// SIMATIC S7-200 project (STEP 7-Micro/WIN), CPU 226 CN REL 02.01

SYMBOL_TABLE USUARIO1
ANTI_HORARIO     Q0.4     // Giro del brazo en sentido antihorario
HORARIO          Q0.5     // Giro del brazo en sentido horario
CIL_DOBLE        Q0.6     // Extencion del brazo neumatico
ELEVACION        Q0.3     // Elevacion del brazo neumatico
PINZA_ABIERTA    Q1.0     // Pinza abierta del brazo neumatico
PINZA_CERRADA    Q0.7     // Pinza cerrada del brazo neumatico
DIRECCION_MOTOR  Q0.1     // Drceccion del motor (adelante o atras)
HL1              Q1.5     // Lampara de señalizacion amarilla
HL2              Q1.6     // Lampara de señaliacion verde
HL3              Q1.7     // Lampara de señalizacion roja
CIL_ABAJO        I0.3     // Sensor indicador de cilindro abajo
CIL_ARRIBA       I0.4     // Sensor indicador de cilindro arriba
CIL_EXT          I0.7     // Sensor indicador de cilindro doble extendido
CIL_RET          I1.0     // Sensor indicador de cilindro doble retraido
PINZA_CERRADO    I1.1     // Sensor indicador de Pinza cerrada
ROT_DER          I0.6     // Sensor indicador de cilindro rotatorio a la derecha
ROT_IZQ          I0.5     // Sensor indicador de cilindro rotatorio a la izquierda
FIN_CARRERA_IZQ  I0.2     // Final de carrera izquierda
FIN_CARRERA_DER  I0.1     // Final de carrera derecha
INDUCTIVO        I0.0     // Sensor inductivo
E0               M0.0     // Estado 0
E0a              M1.4     // Estado 0a
E1               M0.1     // Estado 1
E2               M0.2     // Estado 2
E3               M0.3     // Estado 3
E4               M0.4     // Estado 4
E5               M0.5     // Estaro 5
E6               M0.6     // Estado 6
E7               M0.7     // Estado 7
E8               M1.0     // Estado 8
E9               M1.1     // Estado 9
S1               M1.2     // Estado S1
S2               M1.3     // Estado S2
SBB1             I2.5     // Pulsador de marcha
SBB2             I2.4     // Pulsador de paro
SA               I2.7     // Selector rotativo
QS               I2.6     // Zeta de emergencia
FIN_MOV_1        V50.0    // Posicion de memoria para almacenar el movimiento lineal del brazo neumatico 1
FIN_MOV_2        V50.1    // Posicion de memoria para almacenar el movimiento lineal del brazo neumatico 2
FIN_MOV_3        V50.2    // Posicion de memoria para almacenar el movimiento lineal del brazo neumatico 3
FIN_MOV_4        V50.3    // Posicion de memoria para almacenar el movimiento lineal del brazo neumatico 4
FIN_MOV_5        V50.4    // Posicion de memoria para almacenar el movimiento lineal del brazo neumatico 5
FIN_MOV_6        V50.5    // Posicion de memoria para almacenar el movimiento lineal del brazo neumatico 6
FIN_MOV_7        V50.6    // Posicion de memoria para almacenar el movimiento lineal del brazo neumatico 7
EA               M1.5     // Estado EA
M1               M1.6     // Estado M1
M2               M1.7     // Estado M2
M3               M2.0     // Estado M3
M4               M2.1     // Estado M4
M5               M2.2     // Estado M5
SAA              M2.3     // Estado SAA
EB               M2.4     // Estado EB
M6               M2.5     // Estado M6
M7               M2.6     // Estado M7
M8               M2.7     // Estado M8
M9               M3.0     // Estado M9
M10              M3.1     // Estado M10
M11              M3.2     // Estado M11
M12              M3.3     // Estado M12
M13              M3.4     // Estado M13
M14              M3.5     // Estado M14
M15              M3.6     // Estado M15
M16              M3.7     // Estado M16
M17              M4.0     // Estado M17
SB               M4.1     // Estado SB
EC               M4.2     // Estado EC
M18              M4.3     // Estado M18
M19              M4.4     // Estado M19
M20              M4.5     // Estado M20
M21              M4.6     // Estado M21
M22              M4.7     // Estado M22
M23              M5.0     // Estado M23
M24              M5.1     // Estado M24
M25              M5.2     // Estado M25
M26              M5.3     // Estado M26
M27              M5.4     // Estado M27
M28              M5.5     // Estado M28
M29              M5.6     // Estado M29
SC               M5.7     // Estado SC
E_D              M6.0     // Estado E_D
M30              M6.1     // Estado M30
M31              M6.2     // Estado M31
M32              M6.3     // Estado M32
M33              M6.4     // Estado M33
SD               M6.5     // Estado SD
ciclo            M7.0     // Bit de indicacion para la comunicacion
error_comunica   M7.1     // Bit indicador si hay error en la comunicacion
GO_ALIMENTACION  V0.0     // Iniciar la unidad de alimentacion desde la unidad de transporte
GO_ENSAMBLAJE    V0.2     // Iniciar la unidad de ensamblaje desde la unidad de transporte
GO_PROCESAMIENTO V0.4     // Iniciar la unidad de procesamiento desde la unidad de transporte
GO_SELECCION     V0.6     // Iniciar la unidad de seleccion desde la unidad de transporte
FIN_ALIMENTACION V1.1     // Indica la finalizacion de la unidad y asi el brazo recoja los cilindros
FIN_ENSAMBLAJE   V2.3     // Indica la finalizacion de la unidad y asi el brazo recoja los cilindros
FIN_PROCESAMIENTO V3.5     // Indica la finalizacion de la unidad y asi el brazo recoja los cilindros
EE1              M7.2     // Estado EE1
EE2              M7.3     // Estado EE2
EE3              M7.4     // Estado EE3
MMA              M7.5     // Estado MMA
EEE              M7.6     // Estado EEE
END_SYMBOL_TABLE

ORGANIZATION_BLOCK PRINCIPAL:OB1
TITLE=COMENTARIOS DEL PROGRAMA
BEGIN
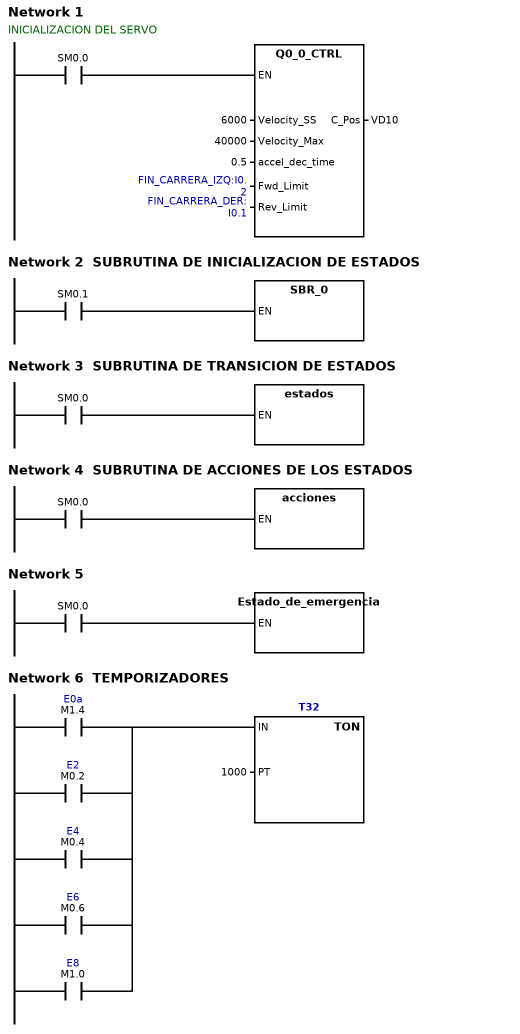
Network 1
// INICIALIZACION DEL SERVO
LD     SM0.0
CALL   Q0_0_CTRL:SBR1, 6000, 40000, 0.5, FIN_CARRERA_IZQ:I0.2, FIN_CARRERA_DER:I0.1, VD10
Network 2 // SUBRUTINA DE INICIALIZACION DE ESTADOS
LD     SM0.1
CALL   SBR_0:SBR0
Network 3 // SUBRUTINA DE TRANSICION DE ESTADOS
LD     SM0.0
CALL   estados:SBR8
Network 4 // SUBRUTINA DE ACCIONES DE LOS ESTADOS
LD     SM0.0
CALL   acciones:SBR9
Network 5
LD     SM0.0
CALL   Estado_de_emergencia:SBR10
Network 6 // TEMPORIZADORES
LD     E0a:M1.4
O      E2:M0.2
O      E4:M0.4
O      E6:M0.6
O      E8:M1.0
TON    T32, 1000
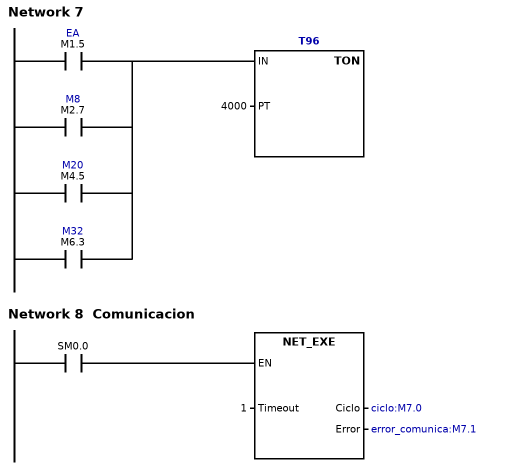
Network 7
LD     EA:M1.5
O      M8:M2.7
O      M20:M4.5
O      M32:M6.3
TON    T96, 4000
Network 8 // Comunicacion	
LD     SM0.0
CALL   NET_EXE:SBR7, 1, ciclo:M7.0, error_comunica:M7.1
END_ORGANIZATION_BLOCK

SUBROUTINE_BLOCK SBR_0:SBR0
TITLE=COMENTARIOS DE LA SUBRUTINA
BEGIN
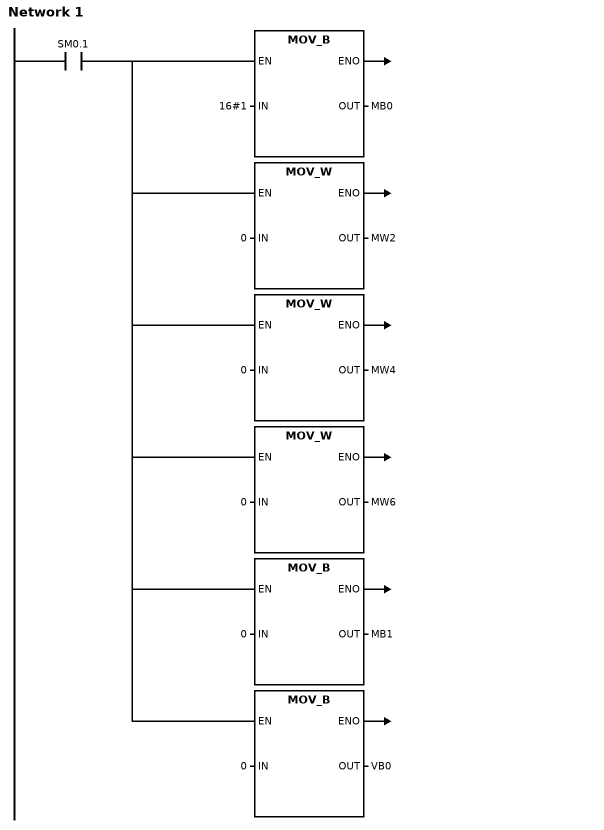
Network 1
LD     SM0.1
MOVB   16#1, MB0
MOVW   0, MW2
MOVW   0, MW4
MOVW   0, MW6
MOVB   0, MB1
MOVB   0, VB0
Network 2 // Título de segmento
// Comentario de segmento
END_SUBROUTINE_BLOCK

// SBR1: protected block, not included

// SBR2: protected block, not included

// SBR3: protected block, not included

// SBR4: protected block, not included

// SBR5: protected block, not included

// SBR6: protected block, not included

// SBR7: protected block, not included

SUBROUTINE_BLOCK estados:SBR8
TITLE=TRANSICION DE ESTADOS
BEGIN
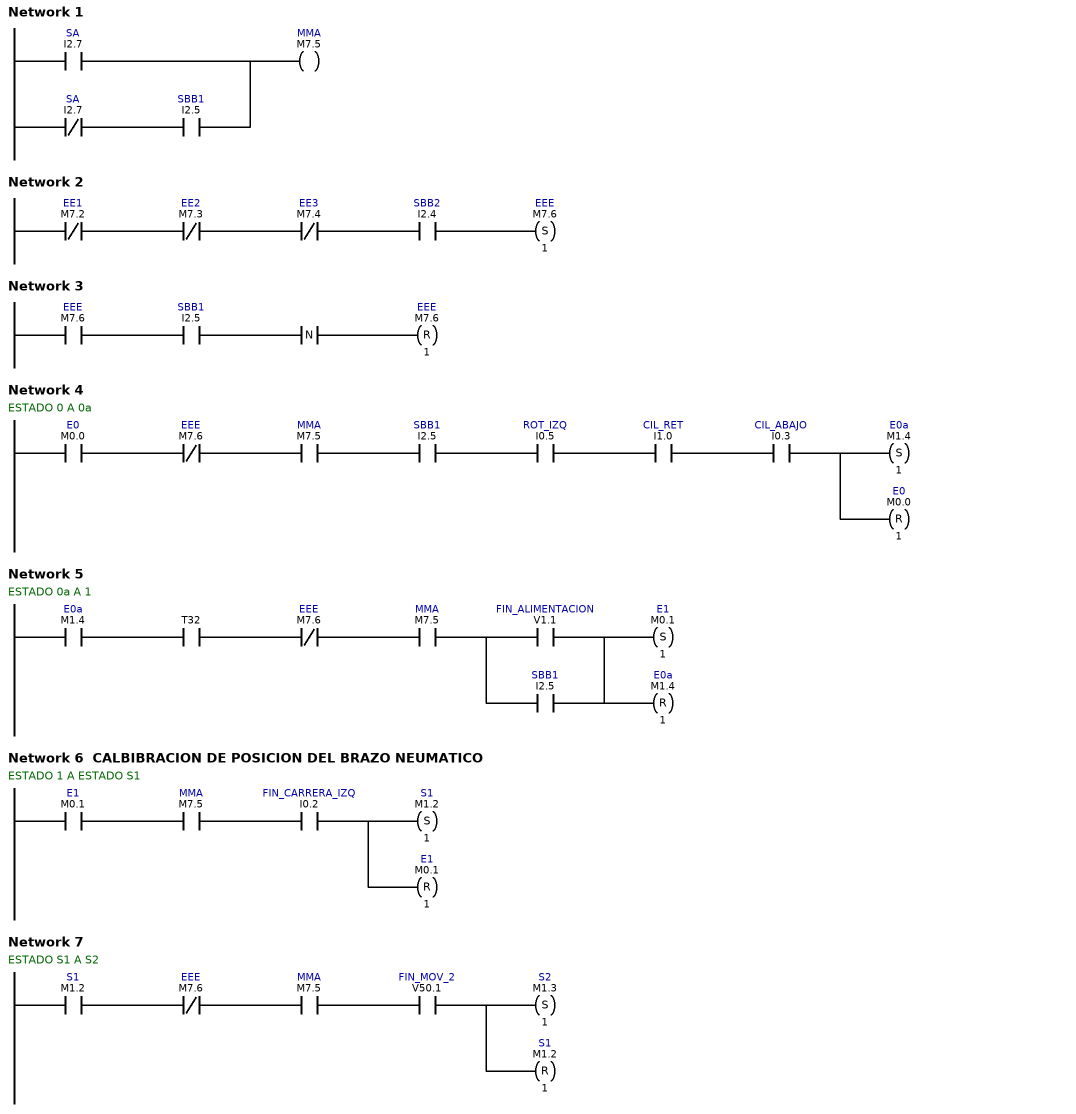
Network 1
LD     SA:I2.7
LDN    SA:I2.7
A      SBB1:I2.5
OLD
=      MMA:M7.5
Network 2
LDN    EE1:M7.2
AN     EE2:M7.3
AN     EE3:M7.4
A      SBB2:I2.4
S      EEE:M7.6, 1
Network 3
LD     EEE:M7.6
A      SBB1:I2.5
ED
R      EEE:M7.6, 1
Network 4
// ESTADO 0 A 0a
LD     E0:M0.0
AN     EEE:M7.6
A      MMA:M7.5
A      SBB1:I2.5
A      ROT_IZQ:I0.5
A      CIL_RET:I1.0
A      CIL_ABAJO:I0.3
S      E0a:M1.4, 1
R      E0:M0.0, 1
Network 5
// ESTADO 0a A 1
LD     E0a:M1.4
A      T32
AN     EEE:M7.6
A      MMA:M7.5
LD     FIN_ALIMENTACION:V1.1
O      SBB1:I2.5
ALD
S      E1:M0.1, 1
R      E0a:M1.4, 1
Network 6 // CALBIBRACION DE POSICION DEL BRAZO NEUMATICO
// ESTADO 1 A ESTADO S1
LD     E1:M0.1
A      MMA:M7.5
A      FIN_CARRERA_IZQ:I0.2
S      S1:M1.2, 1
R      E1:M0.1, 1
Network 7
// ESTADO S1 A S2
LD     S1:M1.2
AN     EEE:M7.6
A      MMA:M7.5
A      FIN_MOV_2:V50.1
S      S2:M1.3, 1
R      S1:M1.2, 1
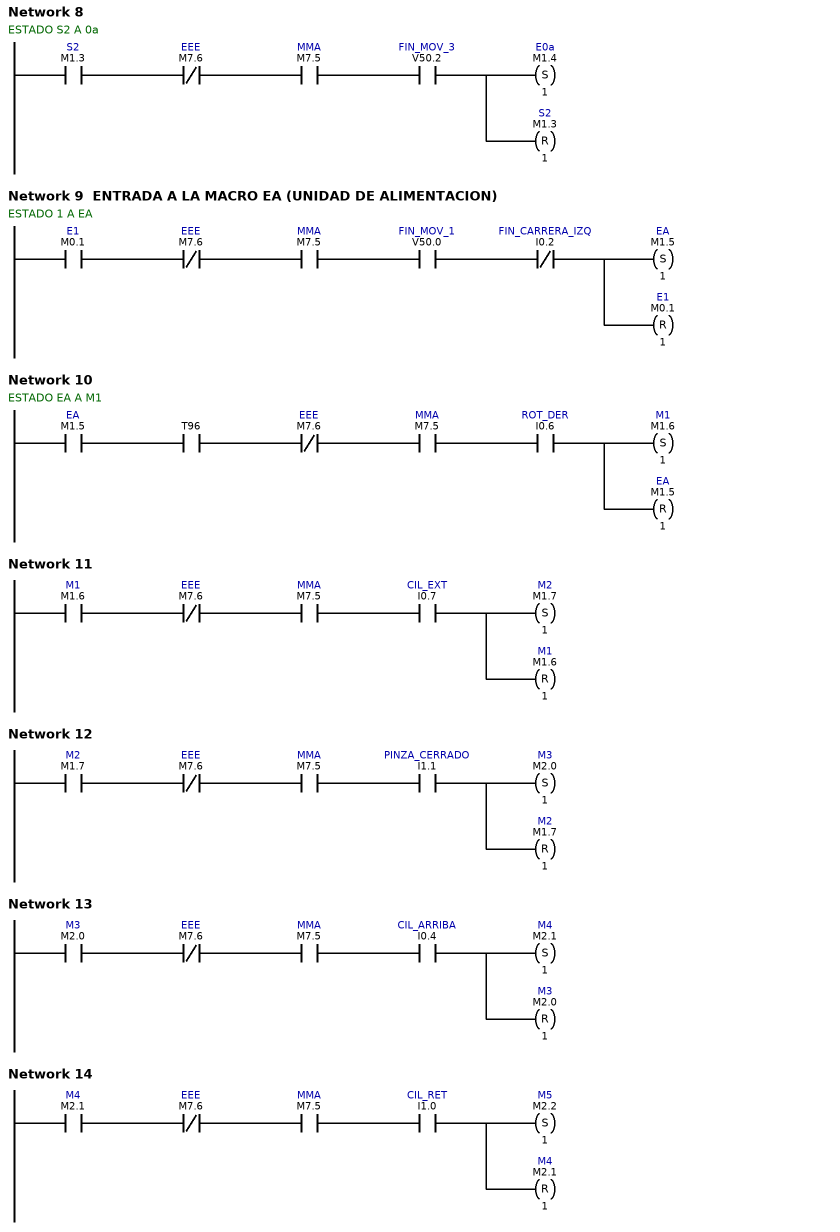
Network 8
// ESTADO S2 A 0a
LD     S2:M1.3
AN     EEE:M7.6
A      MMA:M7.5
A      FIN_MOV_3:V50.2
S      E0a:M1.4, 1
R      S2:M1.3, 1
Network 9 // ENTRADA A LA MACRO EA (UNIDAD DE ALIMENTACION)
// ESTADO 1 A EA
LD     E1:M0.1
AN     EEE:M7.6
A      MMA:M7.5
A      FIN_MOV_1:V50.0
AN     FIN_CARRERA_IZQ:I0.2
S      EA:M1.5, 1
R      E1:M0.1, 1
Network 10
// ESTADO EA A M1
LD     EA:M1.5
A      T96
AN     EEE:M7.6
A      MMA:M7.5
A      ROT_DER:I0.6
S      M1:M1.6, 1
R      EA:M1.5, 1
Network 11
LD     M1:M1.6
AN     EEE:M7.6
A      MMA:M7.5
A      CIL_EXT:I0.7
S      M2:M1.7, 1
R      M1:M1.6, 1
Network 12
LD     M2:M1.7
AN     EEE:M7.6
A      MMA:M7.5
A      PINZA_CERRADO:I1.1
S      M3:M2.0, 1
R      M2:M1.7, 1
Network 13
LD     M3:M2.0
AN     EEE:M7.6
A      MMA:M7.5
A      CIL_ARRIBA:I0.4
S      M4:M2.1, 1
R      M3:M2.0, 1
Network 14
LD     M4:M2.1
AN     EEE:M7.6
A      MMA:M7.5
A      CIL_RET:I1.0
S      M5:M2.2, 1
R      M4:M2.1, 1
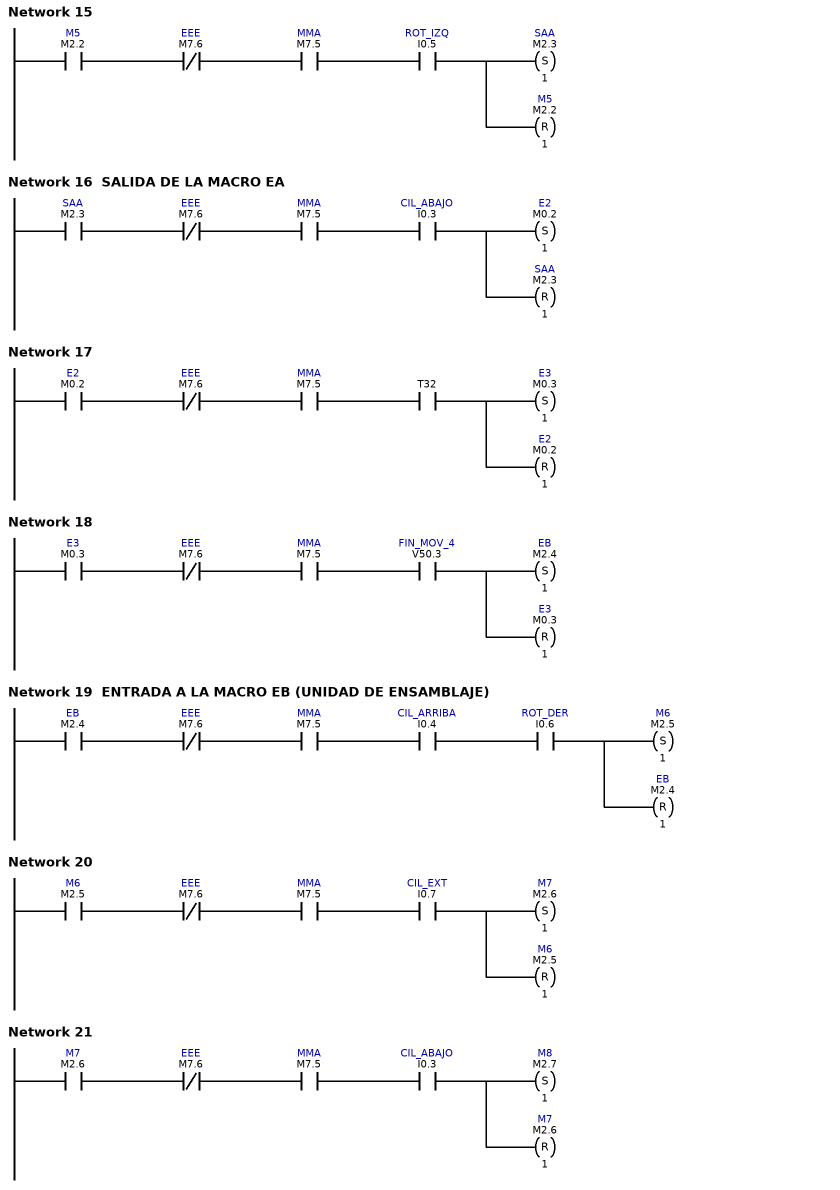
Network 15
LD     M5:M2.2
AN     EEE:M7.6
A      MMA:M7.5
A      ROT_IZQ:I0.5
S      SAA:M2.3, 1
R      M5:M2.2, 1
Network 16 // SALIDA DE LA MACRO EA
LD     SAA:M2.3
AN     EEE:M7.6
A      MMA:M7.5
A      CIL_ABAJO:I0.3
S      E2:M0.2, 1
R      SAA:M2.3, 1
Network 17
LD     E2:M0.2
AN     EEE:M7.6
A      MMA:M7.5
A      T32
S      E3:M0.3, 1
R      E2:M0.2, 1
Network 18
LD     E3:M0.3
AN     EEE:M7.6
A      MMA:M7.5
A      FIN_MOV_4:V50.3
S      EB:M2.4, 1
R      E3:M0.3, 1
Network 19 // ENTRADA A LA MACRO EB (UNIDAD DE ENSAMBLAJE)
LD     EB:M2.4
AN     EEE:M7.6
A      MMA:M7.5
A      CIL_ARRIBA:I0.4
A      ROT_DER:I0.6
S      M6:M2.5, 1
R      EB:M2.4, 1
Network 20
LD     M6:M2.5
AN     EEE:M7.6
A      MMA:M7.5
A      CIL_EXT:I0.7
S      M7:M2.6, 1
R      M6:M2.5, 1
Network 21
LD     M7:M2.6
AN     EEE:M7.6
A      MMA:M7.5
A      CIL_ABAJO:I0.3
S      M8:M2.7, 1
R      M7:M2.6, 1
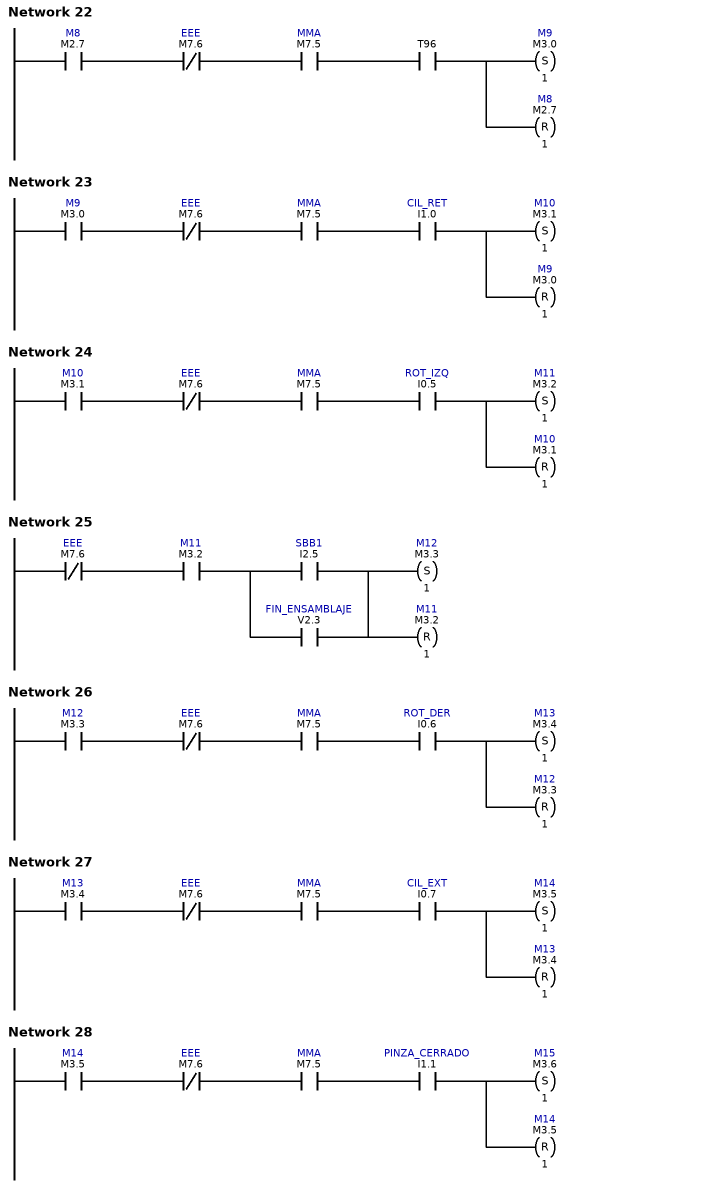
Network 22
LD     M8:M2.7
AN     EEE:M7.6
A      MMA:M7.5
A      T96
S      M9:M3.0, 1
R      M8:M2.7, 1
Network 23
LD     M9:M3.0
AN     EEE:M7.6
A      MMA:M7.5
A      CIL_RET:I1.0
S      M10:M3.1, 1
R      M9:M3.0, 1
Network 24
LD     M10:M3.1
AN     EEE:M7.6
A      MMA:M7.5
A      ROT_IZQ:I0.5
S      M11:M3.2, 1
R      M10:M3.1, 1
Network 25
LDN    EEE:M7.6
A      M11:M3.2
LD     SBB1:I2.5
O      FIN_ENSAMBLAJE:V2.3
ALD
S      M12:M3.3, 1
R      M11:M3.2, 1
Network 26
LD     M12:M3.3
AN     EEE:M7.6
A      MMA:M7.5
A      ROT_DER:I0.6
S      M13:M3.4, 1
R      M12:M3.3, 1
Network 27
LD     M13:M3.4
AN     EEE:M7.6
A      MMA:M7.5
A      CIL_EXT:I0.7
S      M14:M3.5, 1
R      M13:M3.4, 1
Network 28
LD     M14:M3.5
AN     EEE:M7.6
A      MMA:M7.5
A      PINZA_CERRADO:I1.1
S      M15:M3.6, 1
R      M14:M3.5, 1
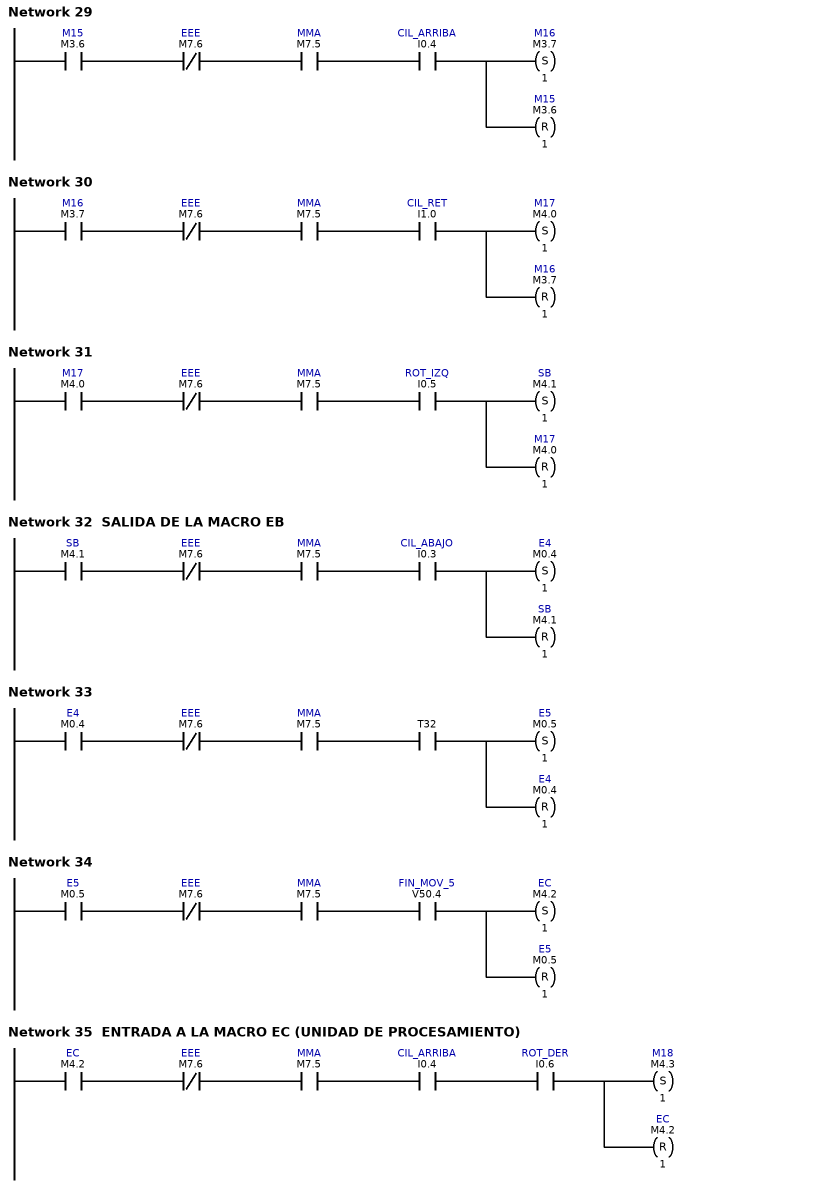
Network 29
LD     M15:M3.6
AN     EEE:M7.6
A      MMA:M7.5
A      CIL_ARRIBA:I0.4
S      M16:M3.7, 1
R      M15:M3.6, 1
Network 30
LD     M16:M3.7
AN     EEE:M7.6
A      MMA:M7.5
A      CIL_RET:I1.0
S      M17:M4.0, 1
R      M16:M3.7, 1
Network 31
LD     M17:M4.0
AN     EEE:M7.6
A      MMA:M7.5
A      ROT_IZQ:I0.5
S      SB:M4.1, 1
R      M17:M4.0, 1
Network 32 // SALIDA DE LA MACRO EB
LD     SB:M4.1
AN     EEE:M7.6
A      MMA:M7.5
A      CIL_ABAJO:I0.3
S      E4:M0.4, 1
R      SB:M4.1, 1
Network 33
LD     E4:M0.4
AN     EEE:M7.6
A      MMA:M7.5
A      T32
S      E5:M0.5, 1
R      E4:M0.4, 1
Network 34
LD     E5:M0.5
AN     EEE:M7.6
A      MMA:M7.5
A      FIN_MOV_5:V50.4
S      EC:M4.2, 1
R      E5:M0.5, 1
Network 35 // ENTRADA A LA MACRO EC (UNIDAD DE PROCESAMIENTO)
LD     EC:M4.2
AN     EEE:M7.6
A      MMA:M7.5
A      CIL_ARRIBA:I0.4
A      ROT_DER:I0.6
S      M18:M4.3, 1
R      EC:M4.2, 1
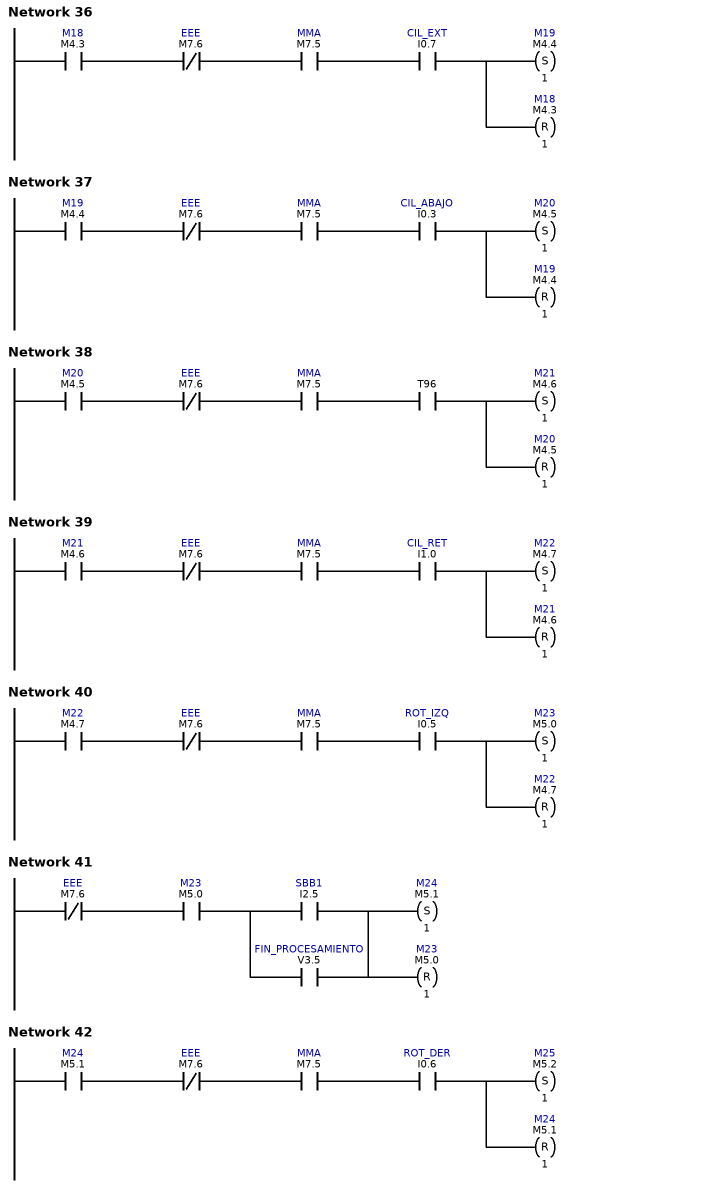
Network 36
LD     M18:M4.3
AN     EEE:M7.6
A      MMA:M7.5
A      CIL_EXT:I0.7
S      M19:M4.4, 1
R      M18:M4.3, 1
Network 37
LD     M19:M4.4
AN     EEE:M7.6
A      MMA:M7.5
A      CIL_ABAJO:I0.3
S      M20:M4.5, 1
R      M19:M4.4, 1
Network 38
LD     M20:M4.5
AN     EEE:M7.6
A      MMA:M7.5
A      T96
S      M21:M4.6, 1
R      M20:M4.5, 1
Network 39
LD     M21:M4.6
AN     EEE:M7.6
A      MMA:M7.5
A      CIL_RET:I1.0
S      M22:M4.7, 1
R      M21:M4.6, 1
Network 40
LD     M22:M4.7
AN     EEE:M7.6
A      MMA:M7.5
A      ROT_IZQ:I0.5
S      M23:M5.0, 1
R      M22:M4.7, 1
Network 41
LDN    EEE:M7.6
A      M23:M5.0
LD     SBB1:I2.5
O      FIN_PROCESAMIENTO:V3.5
ALD
S      M24:M5.1, 1
R      M23:M5.0, 1
Network 42
LD     M24:M5.1
AN     EEE:M7.6
A      MMA:M7.5
A      ROT_DER:I0.6
S      M25:M5.2, 1
R      M24:M5.1, 1
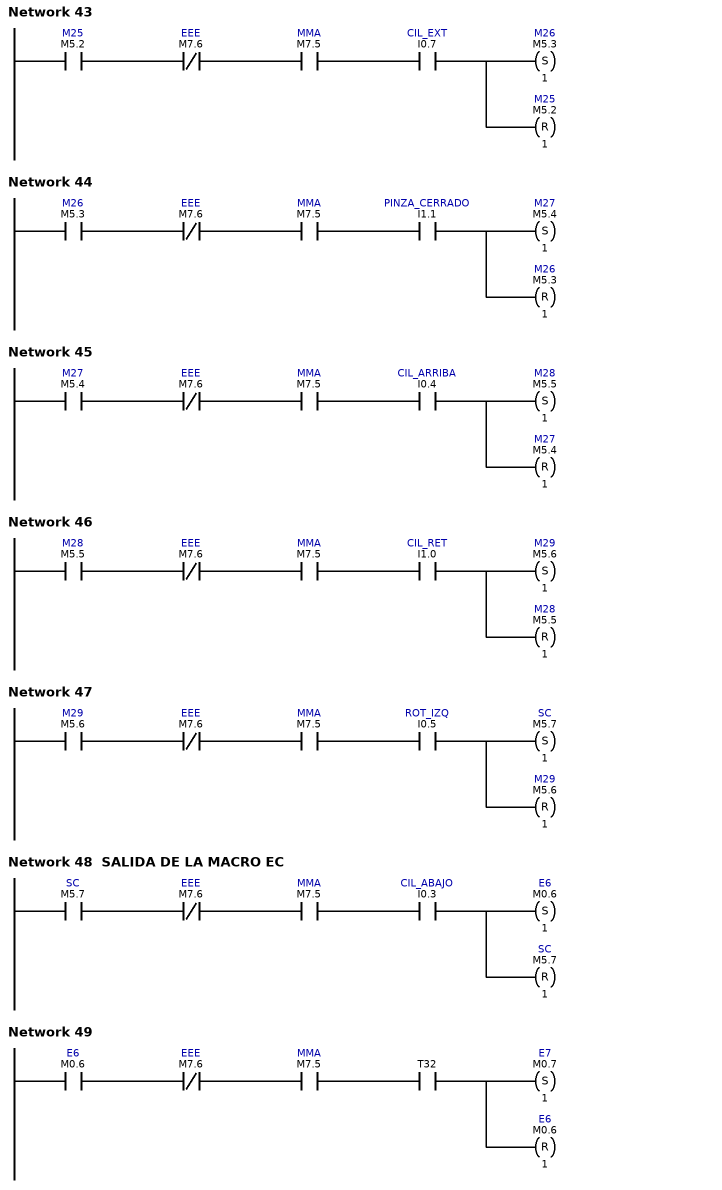
Network 43
LD     M25:M5.2
AN     EEE:M7.6
A      MMA:M7.5
A      CIL_EXT:I0.7
S      M26:M5.3, 1
R      M25:M5.2, 1
Network 44
LD     M26:M5.3
AN     EEE:M7.6
A      MMA:M7.5
A      PINZA_CERRADO:I1.1
S      M27:M5.4, 1
R      M26:M5.3, 1
Network 45
LD     M27:M5.4
AN     EEE:M7.6
A      MMA:M7.5
A      CIL_ARRIBA:I0.4
S      M28:M5.5, 1
R      M27:M5.4, 1
Network 46
LD     M28:M5.5
AN     EEE:M7.6
A      MMA:M7.5
A      CIL_RET:I1.0
S      M29:M5.6, 1
R      M28:M5.5, 1
Network 47
LD     M29:M5.6
AN     EEE:M7.6
A      MMA:M7.5
A      ROT_IZQ:I0.5
S      SC:M5.7, 1
R      M29:M5.6, 1
Network 48 // SALIDA DE LA MACRO EC
LD     SC:M5.7
AN     EEE:M7.6
A      MMA:M7.5
A      CIL_ABAJO:I0.3
S      E6:M0.6, 1
R      SC:M5.7, 1
Network 49
LD     E6:M0.6
AN     EEE:M7.6
A      MMA:M7.5
A      T32
S      E7:M0.7, 1
R      E6:M0.6, 1
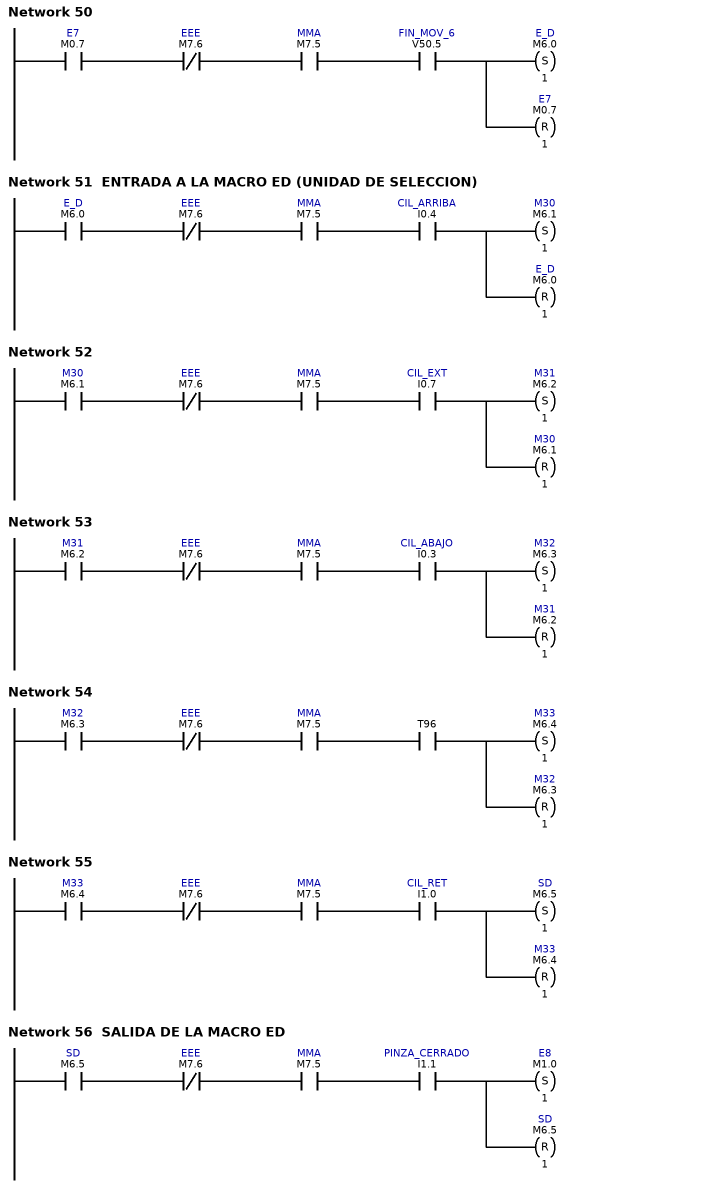
Network 50
LD     E7:M0.7
AN     EEE:M7.6
A      MMA:M7.5
A      FIN_MOV_6:V50.5
S      E_D:M6.0, 1
R      E7:M0.7, 1
Network 51 // ENTRADA A LA MACRO ED (UNIDAD DE SELECCION)
LD     E_D:M6.0
AN     EEE:M7.6
A      MMA:M7.5
A      CIL_ARRIBA:I0.4
S      M30:M6.1, 1
R      E_D:M6.0, 1
Network 52
LD     M30:M6.1
AN     EEE:M7.6
A      MMA:M7.5
A      CIL_EXT:I0.7
S      M31:M6.2, 1
R      M30:M6.1, 1
Network 53
LD     M31:M6.2
AN     EEE:M7.6
A      MMA:M7.5
A      CIL_ABAJO:I0.3
S      M32:M6.3, 1
R      M31:M6.2, 1
Network 54
LD     M32:M6.3
AN     EEE:M7.6
A      MMA:M7.5
A      T96
S      M33:M6.4, 1
R      M32:M6.3, 1
Network 55
LD     M33:M6.4
AN     EEE:M7.6
A      MMA:M7.5
A      CIL_RET:I1.0
S      SD:M6.5, 1
R      M33:M6.4, 1
Network 56 // SALIDA DE LA MACRO ED
LD     SD:M6.5
AN     EEE:M7.6
A      MMA:M7.5
A      PINZA_CERRADO:I1.1
S      E8:M1.0, 1
R      SD:M6.5, 1
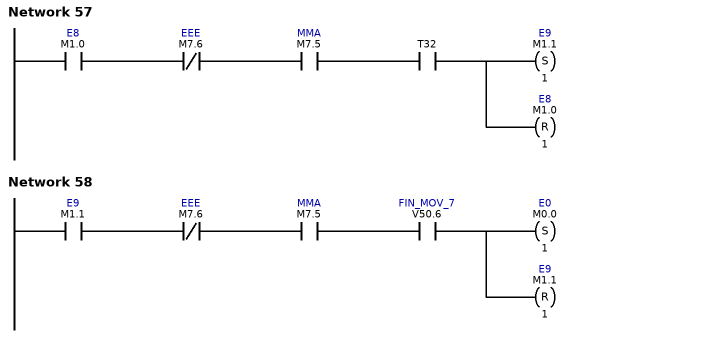
Network 57
LD     E8:M1.0
AN     EEE:M7.6
A      MMA:M7.5
A      T32
S      E9:M1.1, 1
R      E8:M1.0, 1
Network 58
LD     E9:M1.1
AN     EEE:M7.6
A      MMA:M7.5
A      FIN_MOV_7:V50.6
S      E0:M0.0, 1
R      E9:M1.1, 1
END_SUBROUTINE_BLOCK

SUBROUTINE_BLOCK acciones:SBR9
TITLE=ACCIONES
BEGIN
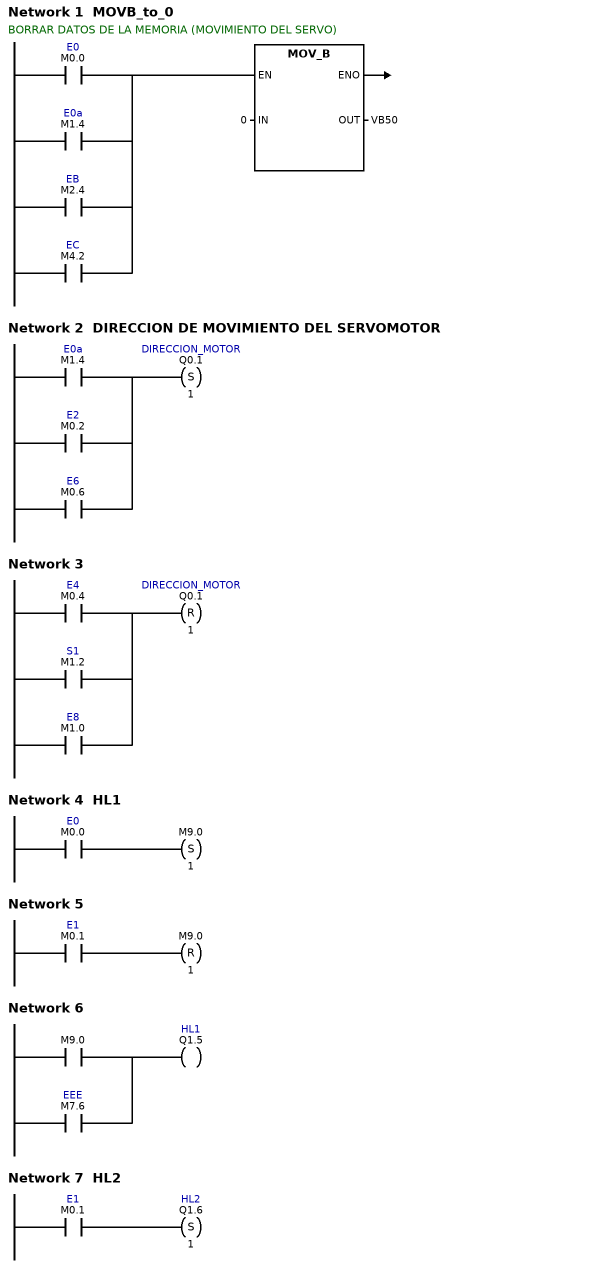
Network 1 // MOVB_to_0
// BORRAR DATOS DE LA MEMORIA (MOVIMIENTO DEL SERVO)
LD     E0:M0.0
O      E0a:M1.4
O      EB:M2.4
O      EC:M4.2
MOVB   0, VB50
Network 2 // DIRECCION DE MOVIMIENTO DEL SERVOMOTOR
LD     E0a:M1.4
O      E2:M0.2
O      E6:M0.6
S      DIRECCION_MOTOR:Q0.1, 1
Network 3
LD     E4:M0.4
O      S1:M1.2
O      E8:M1.0
R      DIRECCION_MOTOR:Q0.1, 1
Network 4 // HL1
LD     E0:M0.0
S      M9.0, 1
Network 5
LD     E1:M0.1
R      M9.0, 1
Network 6
LD     M9.0
O      EEE:M7.6
=      HL1:Q1.5
Network 7 // HL2
LD     E1:M0.1
S      HL2:Q1.6, 1
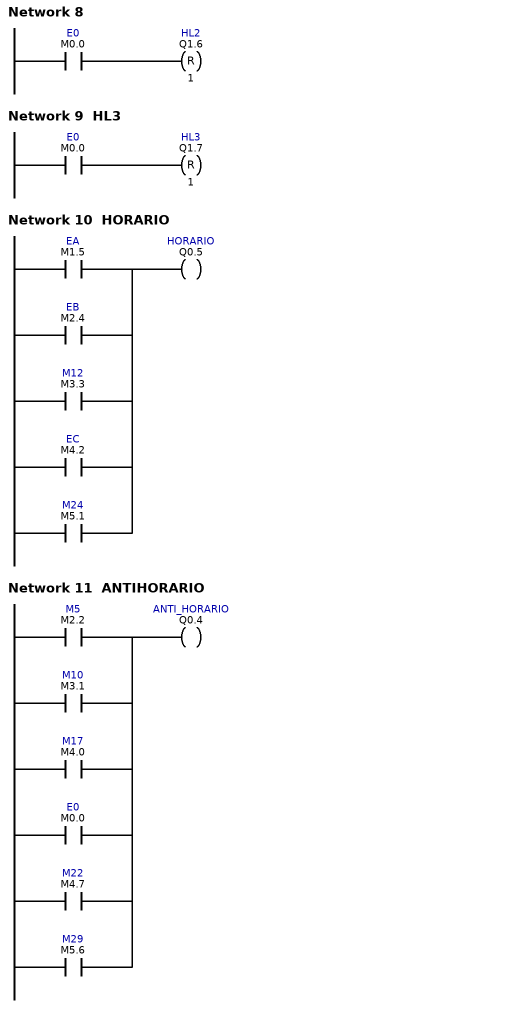
Network 8
LD     E0:M0.0
R      HL2:Q1.6, 1
Network 9 // HL3
LD     E0:M0.0
R      HL3:Q1.7, 1
Network 10 // HORARIO
LD     EA:M1.5
O      EB:M2.4
O      M12:M3.3
O      EC:M4.2
O      M24:M5.1
=      HORARIO:Q0.5
Network 11 // ANTIHORARIO
LD     M5:M2.2
O      M10:M3.1
O      M17:M4.0
O      E0:M0.0
O      M22:M4.7
O      M29:M5.6
=      ANTI_HORARIO:Q0.4
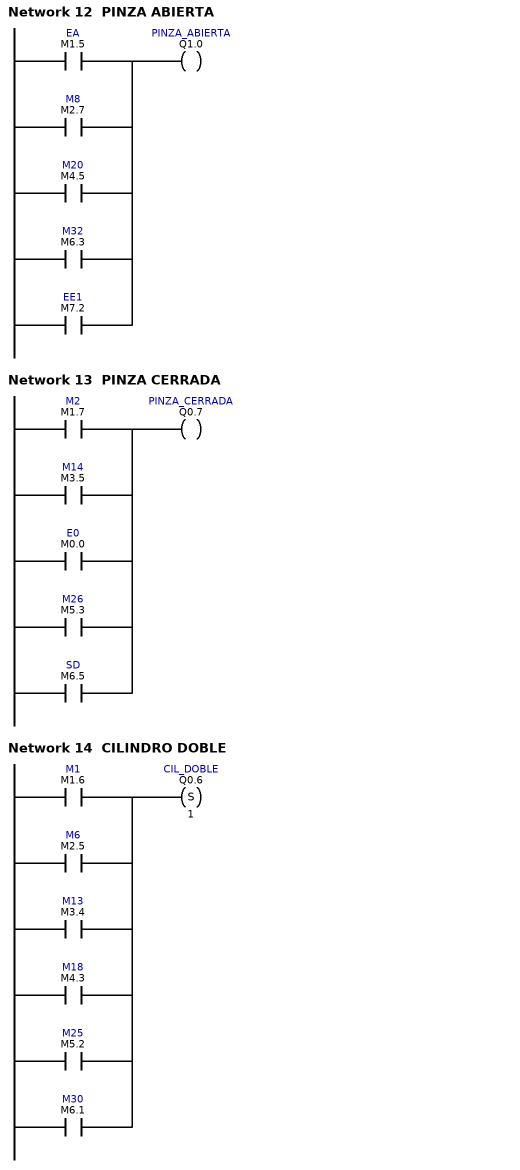
Network 12 // PINZA ABIERTA
LD     EA:M1.5
O      M8:M2.7
O      M20:M4.5
O      M32:M6.3
O      EE1:M7.2
=      PINZA_ABIERTA:Q1.0
Network 13 // PINZA CERRADA
LD     M2:M1.7
O      M14:M3.5
O      E0:M0.0
O      M26:M5.3
O      SD:M6.5
=      PINZA_CERRADA:Q0.7
Network 14 // CILINDRO DOBLE
LD     M1:M1.6
O      M6:M2.5
O      M13:M3.4
O      M18:M4.3
O      M25:M5.2
O      M30:M6.1
S      CIL_DOBLE:Q0.6, 1
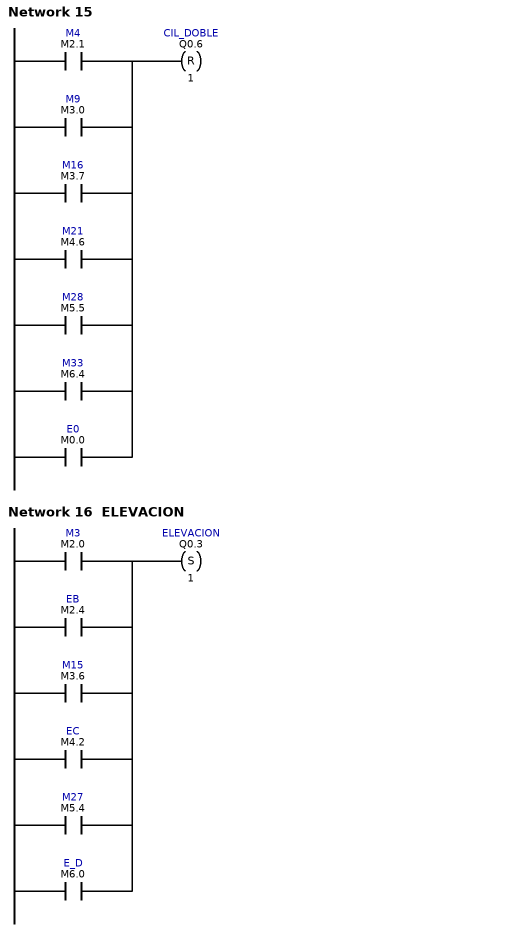
Network 15
LD     M4:M2.1
O      M9:M3.0
O      M16:M3.7
O      M21:M4.6
O      M28:M5.5
O      M33:M6.4
O      E0:M0.0
R      CIL_DOBLE:Q0.6, 1
Network 16 // ELEVACION
LD     M3:M2.0
O      EB:M2.4
O      M15:M3.6
O      EC:M4.2
O      M27:M5.4
O      E_D:M6.0
S      ELEVACION:Q0.3, 1
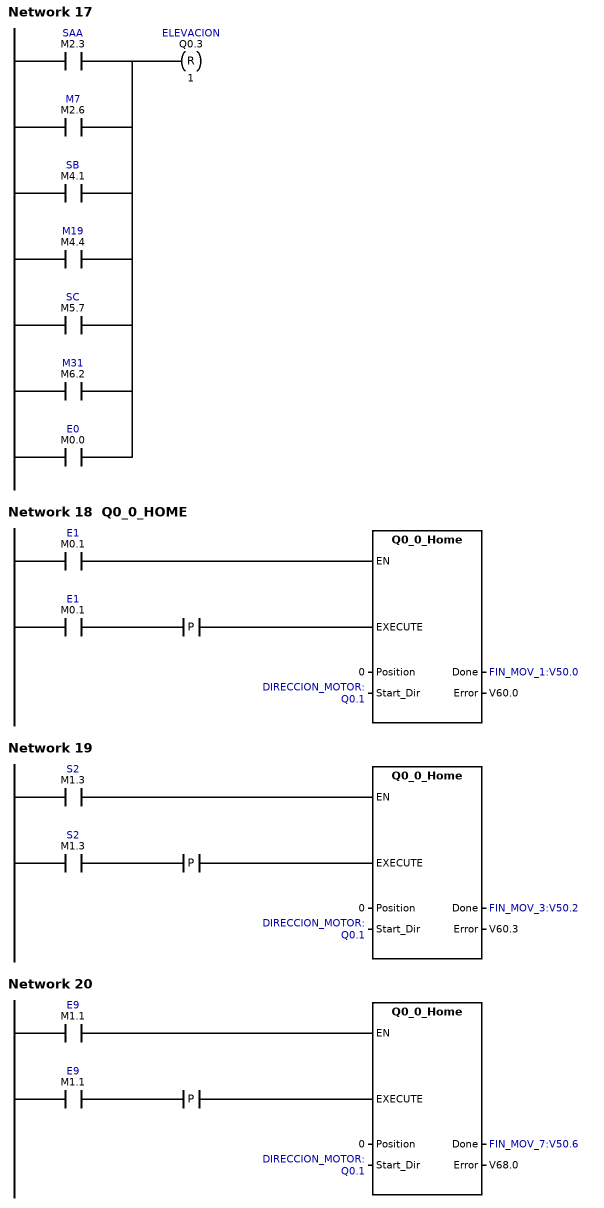
Network 17
LD     SAA:M2.3
O      M7:M2.6
O      SB:M4.1
O      M19:M4.4
O      SC:M5.7
O      M31:M6.2
O      E0:M0.0
R      ELEVACION:Q0.3, 1
Network 18 // Q0_0_HOME
LD     E1:M0.1
=      L60.0
LD     E1:M0.1
EU
=      L63.7
LD     L60.0
CALL   Q0_0_Home:SBR3, L63.7, 0, DIRECCION_MOTOR:Q0.1, FIN_MOV_1:V50.0, V60.0
Network 19
LD     S2:M1.3
=      L60.0
LD     S2:M1.3
EU
=      L63.7
LD     L60.0
CALL   Q0_0_Home:SBR3, L63.7, 0, DIRECCION_MOTOR:Q0.1, FIN_MOV_3:V50.2, V60.3
Network 20
LD     E9:M1.1
=      L60.0
LD     E9:M1.1
EU
=      L63.7
LD     L60.0
CALL   Q0_0_Home:SBR3, L63.7, 0, DIRECCION_MOTOR:Q0.1, FIN_MOV_7:V50.6, V68.0
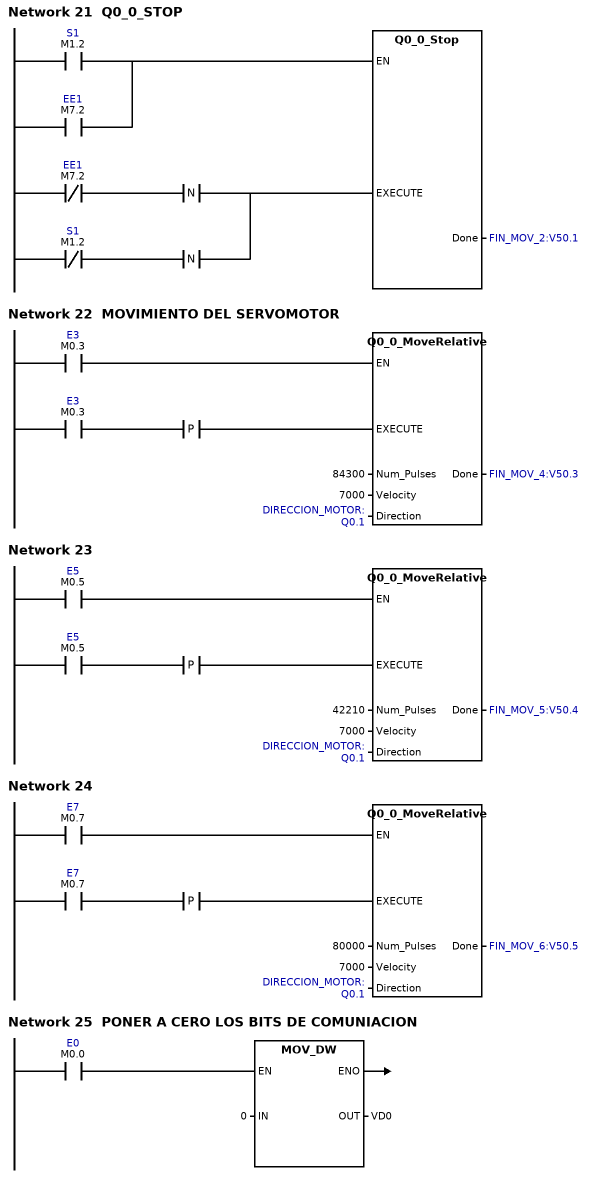
Network 21 // Q0_0_STOP
LD     S1:M1.2
O      EE1:M7.2
=      L60.0
LDN    EE1:M7.2
ED
LDN    S1:M1.2
ED
OLD
=      L63.7
LD     L60.0
CALL   Q0_0_Stop:SBR6, L63.7, FIN_MOV_2:V50.1
Network 22 // MOVIMIENTO DEL SERVOMOTOR
LD     E3:M0.3
=      L60.0
LD     E3:M0.3
EU
=      L63.7
LD     L60.0
CALL   Q0_0_MoveRelative:SBR4, L63.7, 84300, 7000, DIRECCION_MOTOR:Q0.1, FIN_MOV_4:V50.3
Network 23
LD     E5:M0.5
=      L60.0
LD     E5:M0.5
EU
=      L63.7
LD     L60.0
CALL   Q0_0_MoveRelative:SBR4, L63.7, 42210, 7000, DIRECCION_MOTOR:Q0.1, FIN_MOV_5:V50.4
Network 24
LD     E7:M0.7
=      L60.0
LD     E7:M0.7
EU
=      L63.7
LD     L60.0
CALL   Q0_0_MoveRelative:SBR4, L63.7, 80000, 7000, DIRECCION_MOTOR:Q0.1, FIN_MOV_6:V50.5
Network 25 // PONER A CERO LOS BITS DE COMUNIACION
LD     E0:M0.0
MOVD   0, VD0
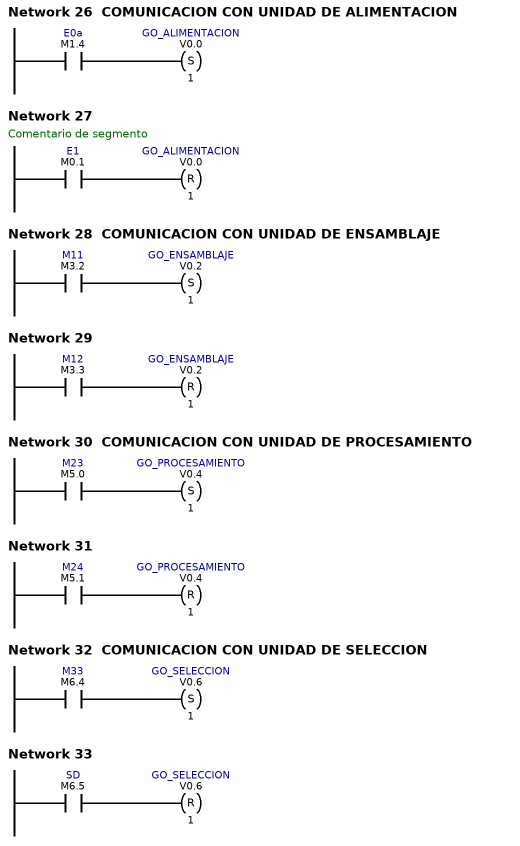
Network 26 // COMUNICACION CON UNIDAD DE ALIMENTACION
LD     E0a:M1.4
S      GO_ALIMENTACION:V0.0, 1
Network 27
// Comentario de segmento
LD     E1:M0.1
R      GO_ALIMENTACION:V0.0, 1
Network 28 // COMUNICACION CON UNIDAD DE ENSAMBLAJE
LD     M11:M3.2
S      GO_ENSAMBLAJE:V0.2, 1
Network 29
LD     M12:M3.3
R      GO_ENSAMBLAJE:V0.2, 1
Network 30 // COMUNICACION CON UNIDAD DE PROCESAMIENTO
LD     M23:M5.0
S      GO_PROCESAMIENTO:V0.4, 1
Network 31
LD     M24:M5.1
R      GO_PROCESAMIENTO:V0.4, 1
Network 32 // COMUNICACION CON UNIDAD DE SELECCION
LD     M33:M6.4
S      GO_SELECCION:V0.6, 1
Network 33
LD     SD:M6.5
R      GO_SELECCION:V0.6, 1
END_SUBROUTINE_BLOCK

SUBROUTINE_BLOCK Estado_de_emergencia:SBR10
TITLE=COMENTARIOS DE LA SUBRUTINA
BEGIN
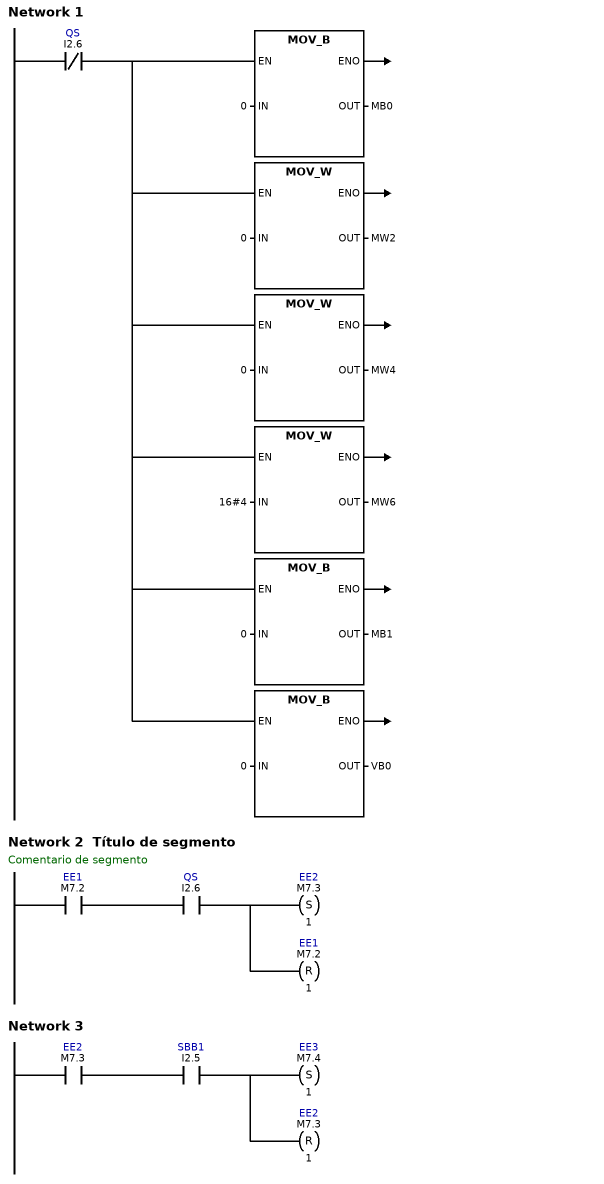
Network 1
LDN    QS:I2.6
MOVB   0, MB0
MOVW   0, MW2
MOVW   0, MW4
MOVW   16#4, MW6
MOVB   0, MB1
MOVB   0, VB0
Network 2 // Título de segmento
// Comentario de segmento
LD     EE1:M7.2
A      QS:I2.6
S      EE2:M7.3, 1
R      EE1:M7.2, 1
Network 3
LD     EE2:M7.3
A      SBB1:I2.5
S      EE3:M7.4, 1
R      EE2:M7.3, 1
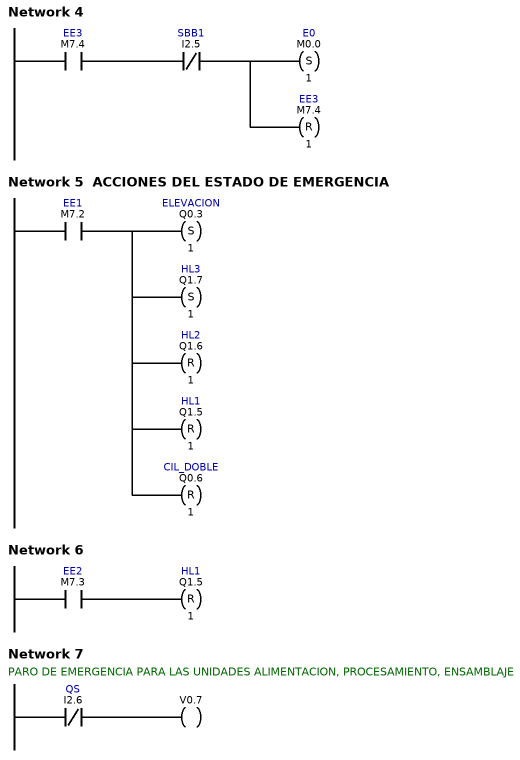
Network 4
LD     EE3:M7.4
AN     SBB1:I2.5
S      E0:M0.0, 1
R      EE3:M7.4, 1
Network 5 // ACCIONES DEL ESTADO DE EMERGENCIA
LD     EE1:M7.2
S      ELEVACION:Q0.3, 1
S      HL3:Q1.7, 1
R      HL2:Q1.6, 1
R      HL1:Q1.5, 1
R      CIL_DOBLE:Q0.6, 1
Network 6
LD     EE2:M7.3
R      HL1:Q1.5, 1
Network 7
// PARO DE EMERGENCIA PARA LAS UNIDADES ALIMENTACION, PROCESAMIENTO, ENSAMBLAJE 
LDN    QS:I2.6
=      V0.7
END_SUBROUTINE_BLOCK
